(*
SPDX-FileCopyrightText: © 2026 Oleksandr Tiutyk <trofimich@gmail.com>
SPDX-License-Identifier: MIT
License: https://opensource.org/license/mit
*)

(*!
<summary>Describes an action by name without executing it or carrying additional action parameters.</summary>
<description>
The initialization name is copied into instance storage and exposed through the read-only INamed contract.
Names are expected to be nonempty, but are not required to be globally unique. Each permission policy defines
how it recognizes an action; equal names alone do not establish action identity.
</description>
*)

{attribute 'no_explicit_call' := 'do not call this function block directly'}
FUNCTION_BLOCK SimpleActionDescriptor EXTENDS Object IMPLEMENTS INamed
VAR_STAT
	//! <summary>Class name shared by all instances of this function block.</summary>
	{attribute 'hide'} 
	_ClassName : STRING := __POUNAME();
END_VAR
VAR
	{attribute 'hide'} 
	_Name : WSTRING;
END_VAR

{attribute 'monitoring' := 'call'}
PROPERTY ClassName : REFERENCE TO STRING
GET
ClassName REF= _ClassName;
END_GET
END_PROPERTY

(*!
<summary>Copies the action name into instance storage.</summary>
<description>
The name must be nonempty under the action descriptor contract. No allocation or exception is performed; input
storage is not retained.
</description>
*)
METHOD FB_init : BOOL
VAR_INPUT
	bInitRetains : BOOL; // TRUE: the retain variables are initialized (reset warm / reset cold)
	bInCopyCode : BOOL;  // TRUE: the instance will be copied to the copy code afterward (online change)
	name : WSTRING;
END_VAR
_Name := name;
END_METHOD

(*!
<summary>Exposes the action name without copying it.</summary>
<description>
Borrowed read-only reference valid for the descriptor lifetime. The name is fixed by initialization and must
not be changed through this reference.
</description>
*)
{attribute 'monitoring' := 'call'}
PROPERTY FINAL Name : REFERENCE TO WSTRING
GET
Name REF= _Name;
END_GET
END_PROPERTY

(*!
<summary>Provides the library namespace used in diagnostics.</summary>
<description>
Borrowed read-only reference to the compiler-initialized library namespace; no ownership transfer.
</description>
*)
{attribute 'monitoring' := 'call'}
PROPERTY NamespaceName : REFERENCE TO STRING
GET
NamespaceName REF= CurrentNamespace.Name;
END_GET
END_PROPERTY

(*!
<summary>Reports the byte size of this concrete instance.</summary>
<description>
Uses XSIZEOF on the instance. Does not include separately allocated payloads or prove that an arbitrary
address is valid.
</description>
*)
{attribute 'monitoring' := 'call'}
PROPERTY SelfSize : ULINT
GET
SelfSize := XSIZEOF(THIS^);
END_GET
END_PROPERTY

END_FUNCTION_BLOCK

(* stored: Version 1.1.0.1
   POU SimpleActionDescriptor: Id {856aea8e-1241-4104-8feb-5476cb8fbca8}, SpecialFunc None
   Property ClassName: Id {3142e366-b89b-4444-b764-3f825bdc6d6a}
   Get Get: Id {b9a94c6b-1edf-4d76-af80-87d37d88f65f}
   Method FB_init: Id {a67d048a-93ef-4047-b96f-e73d16ee7e8e}
   Property Name: Id {03c97eee-32bf-4e2c-9c90-9e076a537e2f}
   Get Get: Id {8b41e209-52ce-40af-95c1-7b332322dbeb}
   Property NamespaceName: Id {263264a5-c98e-41b5-b8bb-05dda72b5bcd}
   Get Get: Id {1c29f2f5-90c5-4a3d-9532-19ff96ae710b}
   Property SelfSize: Id {39772ead-cc6e-4411-b576-e0b71a5afce1}
   Get Get: Id {4ab3c840-35da-42e6-8f34-5ae16131d9ce} *)
